       // Update validation flag in DB
       "DB_Recipes".Active_Recipe.Recipe_Valid := #Recipe_Valid;
       #Operation_OK := TRUE;
   END_IF;
END_FUNCTION

FUNCTION "FC_Safety_Monitor" : Void   // FC6, SCL
{ S7_Optimized_Access := 'TRUE' }
VERSION : 0.1
   VAR_INPUT
      Emergency_Stop : Bool;
      Door_Interlock_OK : Bool;
      Door_Locked : Bool;
      Manhole_Secured : Bool;
      Temperature_Value : Real;
      Pressure_Value : Real;
      System_Enabled : Bool;
   END_VAR
   VAR_OUTPUT
      Safety_OK : Bool;
      System_Ready : Bool;
      Emergency_Active : Bool;
      Safety_Fault : Bool;
      Fault_Code : UInt;
      Fault_Text : String;
   END_VAR
   VAR_TEMP
      Temp_High_Limit : Real;
      Pressure_High_Limit : Real;
   END_VAR
BEGIN
   #Safety_OK := TRUE;
   #Safety_Fault := FALSE;
   #Fault_Text := '';
   IF #Emergency_Stop THEN
       #Safety_OK := FALSE;
       #Safety_Fault := TRUE;
       #Fault_Text := 'EMERGENCY STOP ACTIVE';
       #System_Ready := FALSE;
       RETURN;
   END_IF;
   IF NOT #Door_Interlock_OK THEN
       #Safety_OK := FALSE;
       #Safety_Fault := TRUE;
       #Fault_Text := 'Door interlock not OK';
   END_IF;
   IF #Temperature_Value > 105.0 THEN
       #Safety_OK := FALSE;
       #Safety_Fault := TRUE;
       #Fault_Text := 'Temperature too high';
   END_IF;
   IF #Pressure_Value > 2500.0 THEN
       #Safety_OK := FALSE;
       #Safety_Fault := TRUE;
       #Fault_Text := 'Pressure too high';
   END_IF;
   #System_Ready := #Safety_OK AND #System_Enabled;
   IF #Safety_OK THEN
       #Fault_Text := 'All safety systems OK';
   END_IF;
END_FUNCTION

FUNCTION "FC_Lock_Discharge_Door" : Void   // FC7, SCL
{ S7_Optimized_Access := 'TRUE' }
VERSION : 0.1
   VAR_INPUT
      Step_Enable : Bool;
      Safety_OK : Bool;
      Step_Timeout : Time;
      Door_Locked_FB : Bool;
      Reset_Step : Bool;
   END_VAR
   VAR_OUTPUT
      Step_Complete : Bool;
      Step_Active : Bool;
      Step_Fault : Bool;
      Fault_Code : UInt;
      Status_Text : String;   // // Step status description
      Time_Remaining : Time;
   END_VAR
   VAR_IN_OUT
      Step_Timer : TON_TIME;
      Close_Timer : TON_TIME;
   END_VAR
BEGIN
   IF #Reset_Step THEN
       #Step_Timer(IN := FALSE,
                   PT := T#0S);
       #Step_Complete := FALSE;
       #Step_Active := FALSE;
       #Step_Fault := FALSE;
       #Fault_Code := 0;
       #Status_Text := 'Step reset';
       "DB_Valves".Valves[3].Close_Auto := FALSE;      // V3 discharge unlock
       RETURN;
   END_IF;
   IF #Step_Enable AND #Safety_OK THEN
       #Step_Active := TRUE;
       #Status_Text := 'Locking discharge door';

       "DB_Valves".Valves[3].Close_Auto := TRUE;       // V3 discharge unlock - close to
       #Step_Timer(IN := TRUE,
                   PT := #Step_Timeout);
       #Time_Remaining := #Step_Timeout - #Step_Timer.ET;
       #Close_Timer(IN := #Door_Locked_FB,
                    PT := T#2s);



       IF #Close_Timer.Q THEN
           #Step_Complete := TRUE;
           #Step_Active := FALSE;
           #Status_Text := 'Door locked successfully';
           "DB_Valves".Valves[3].Close_Auto := FALSE;

       ELSIF #Step_Timer.Q THEN
           #Step_Complete := FALSE;
           #Step_Active := FALSE;
           #Step_Fault := TRUE;
           #Fault_Code := 15;
           #Status_Text := 'Door lock timeout';
       END_IF;
   ELSE
       #Step_Active := FALSE;
       #Step_Complete := FALSE;
       #Step_Timer(IN := FALSE,
                   PT := T#0S);
       "DB_Valves".Valves[3].Close_Auto := FALSE;
       #Status_Text := 'Step disabled';
   END_IF;
END_FUNCTION

FUNCTION "FC_Add_Water" : Void   // FC8, SCL
{ S7_Optimized_Access := 'TRUE' }
VERSION : 0.1
   VAR_INPUT
      Step_Enable : Bool;
      Safety_OK : Bool;
      Reset_Step : Bool;
      Step_Timeout : Time;
      Target_Quantity : Real;
      Flow_Rate : Real;
   END_VAR
   VAR_OUTPUT
      Step_Complete : Bool;
      Water_Level_FB : Bool;
      Step_Active : Bool;
      Step_Fault : Bool;
      Fault_Code : UInt;
      Status_Text : String;
      Water_Added : Real;
      Time_Remaining : Time;
   END_VAR
   VAR_IN_OUT
      Step_Timer : TON_TIME;
   END_VAR
BEGIN
   IF #Reset_Step THEN
       #Step_Timer(IN := FALSE,
                   PT := T#0S);
       #Step_Complete := FALSE;
       #Step_Active := FALSE;
       #Step_Fault := FALSE;
       #Status_Text := 'Step reset';
       "DB_Valves".Valves[5].Open_Auto := FALSE;       // V5 water
       "DB_Valves".Valves[7].Open_Auto := FALSE;       // V7 evacuation
       #Water_Added := 0.0;
       RETURN;
   END_IF;

   IF #Step_Enable AND #Safety_OK THEN
       #Step_Active := TRUE;
       #Status_Text := 'Adding water';

       "DB_Valves".Valves[5].Open_Auto := TRUE;        // V5 water
       "DB_Valves".Valves[7].Open_Auto := TRUE;        // V7 evacuation
       "DB_Valves".Valves[3].Close_Auto := TRUE;         //V3
       #Step_Timer(IN := TRUE,
                   PT := #Step_Timeout);
       #Time_Remaining := #Step_Timeout - #Step_Timer.ET;

       IF #Flow_Rate > 0.0 THEN
           #Water_Added := (DINT_TO_REAL(TIME_TO_DINT(#Step_Timer.ET)) / 10.0) * #Flow_Rate;
           IF "DB_Recipes".Active_Recipe.Production.Adding_Water1_QTY < #Water_Added THEN
               "DB_Process".IO.Water_Level_FB := TRUE;
           END_IF;
       END_IF;

       IF "DB_Process".IO.Water_Level_FB THEN
           #Step_Complete := TRUE;
           #Step_Active := FALSE;
           #Status_Text := 'Water level reached';
           "DB_Valves".Valves[5].Open_Auto := FALSE;
       ELSIF #Step_Timer.Q THEN
           #Step_Complete := FALSE;
           #Step_Active := FALSE;
           #Step_Fault := TRUE;
           #Fault_Code := 1;
           #Status_Text := 'Water addition timeout';
       END_IF;
   ELSE
       #Step_Active := FALSE;
       #Step_Complete := FALSE;
       #Step_Timer(IN := FALSE,
                   PT := T#0S);
       "DB_Valves".Valves[5].Open_Auto := FALSE;
       "DB_Valves".Valves[7].Open_Auto := FALSE;
       #Status_Text := 'Step disabled';
   END_IF;
END_FUNCTION

FUNCTION "FC_Open_Manhole" : Void   // FC9, SCL
{ S7_Optimized_Access := 'TRUE' }
VERSION : 0.1
   VAR_INPUT
      Step_Enable : Bool;
      Safety_OK : Bool;
      Manhole_Open_FB : Bool;
      Manhole_Closed_FB : Bool;
      Reset_Step : Bool;
      Step_Timeout : Time;
   END_VAR
   VAR_OUTPUT
      Step_Complete : Bool;
      Step_Active : Bool;
      Step_Fault : Bool;
      Fault_Code : UInt;
      Status_Text : String;
      Time_Remaining : Time;   // // Time remaining in step
   END_VAR
   VAR_IN_OUT
      Step_Timer : TON_TIME;
      Open_Timer : TON_TIME;
   END_VAR
BEGIN
   IF #Reset_Step THEN
       #Step_Timer(IN := FALSE,
                   PT := T#0S);
       #Step_Complete := FALSE;
       #Step_Active := FALSE;
       #Step_Fault := FALSE;
       #Status_Text := 'Step reset';
       "DB_Valves".Valves[3].Open_Auto := FALSE;
       "DB_Valves".Valves[1].Open_Auto := FALSE;       // V1 manhole
       RETURN;
   END_IF;
   IF #Step_Enable AND #Safety_OK THEN
       #Step_Active := TRUE;
       #Status_Text := 'Opening manhole';

       "DB_Valves".Valves[1].Open_Auto := TRUE;        // V1 manhole
       "DB_Valves".Valves[3].Open_Auto := TRUE; 
       #Step_Timer(IN := TRUE,
                   PT := #Step_Timeout);
       #Time_Remaining := #Step_Timeout - #Step_Timer.ET;
       #Open_Timer(IN:=#Manhole_Closed_FB,
                   PT:=T#2S);
       IF #Open_Timer.Q THEN
           #Step_Complete := TRUE;
           #Step_Active := FALSE;
           #Status_Text := 'Manhole opened';
       ELSIF #Step_Timer.Q THEN
           #Step_Complete := FALSE;
           #Step_Active := FALSE;
           #Step_Fault := TRUE;
           #Fault_Code := 2;
           #Status_Text := 'Manhole open timeout';
       END_IF;
   ELSE
       #Step_Active := FALSE;
       #Step_Complete := FALSE;
       #Step_Timer(IN := FALSE,
                   PT := T#0S);
       "DB_Valves".Valves[1].Open_Auto := FALSE;
       "DB_Valves".Valves[3].Open_Auto := FALSE;
       #Status_Text := 'Step disabled';
   END_IF;
END_FUNCTION

FUNCTION "FC_Wait_Raw_Materials" : Void   // FC10, SCL
{ S7_Optimized_Access := 'TRUE' }
VERSION : 0.1
   VAR_INPUT
      Step_Enable : Bool;
      Safety_OK : Bool;
      RawMat_Confirm : Bool;   // // Raw materials loaded confirmation
      Manhole_Open_FB : Bool;   // // Manhole open feedback
      Manhole_Closed_FB : Bool;
      Reset_Step : Bool;
      Max_Wait_Time : Time;   // // Maximum wait time
   END_VAR
   VAR_OUTPUT
      Step_Complete : Bool;
      Step_Active : Bool;
      Step_Fault : Bool;
      Fault_Code : UInt;
      Status_Text : String;
      Wait_Time_Elapsed : Time;
   END_VAR
   VAR_IN_OUT
      Wait_Timer : TON_TIME;
   END_VAR
BEGIN
   IF #Reset_Step THEN
       #Wait_Timer(IN := FALSE,
                   PT := T#0S);
       #Step_Complete := FALSE;
       #Step_Active := FALSE;
       #Step_Fault := FALSE;
       #Status_Text := 'Step reset';
       RETURN;
   END_IF;
   IF #Step_Enable AND #Safety_OK THEN
       #Step_Active := TRUE;
       #Status_Text := 'Waiting for raw materials';

       "DB_Valves".Valves[1].Open_Auto := TRUE;        // V1 manhole - keep open
       "DB_Valves".Valves[3].Open_Auto := TRUE;        // V7 evacuation
       #Wait_Timer(IN := TRUE,
                   PT := #Max_Wait_Time);
       #Wait_Time_Elapsed := #Wait_Timer.ET;

       IF  #Manhole_Closed_FB THEN
           #Step_Complete := FALSE;
           #Step_Active := FALSE;
           #Step_Fault := TRUE;
           #Fault_Code := 3;
           #Status_Text := 'Manhole not open-Reset PLS';
           RETURN;
       END_IF;

       IF #RawMat_Confirm THEN
           #Step_Complete := TRUE;
           #Step_Active := FALSE;
           #Status_Text := 'Raw materials confirmed';
       ELSIF #Wait_Timer.Q THEN
           #Status_Text := 'Long wait time - check operator';
           #Wait_Timer(IN := FALSE,
                       PT := T#0S);
       END_IF;
   ELSE
       #Step_Active := FALSE;
       #Step_Complete := FALSE;
       #Wait_Timer(IN := FALSE,
                   PT := T#0S);
       #Status_Text := 'Step disabled';
   END_IF;
END_FUNCTION

FUNCTION "FC_Close_Manhole" : Void   // FC11, SCL
{ S7_Optimized_Access := 'TRUE' }
VERSION : 0.1
   VAR_INPUT
      Step_Enable : Bool;
      Safety_OK : Bool;
      Step_Timeout : Time;
      Manhole_Closed_FB : Bool;
      Reset_Step : Bool;
      Manhole_Open_FB : Bool;
   END_VAR
   VAR_OUTPUT
      Step_Complete : Bool;
      Step_Active : Bool;
      Step_Fault : Bool;
      Fault_Code : UInt;
      Status_Text : String;
      Time_Remaining : Time;
   END_VAR
   VAR_IN_OUT
      Step_Timer : TON_TIME;
      Close_Timer : TON_TIME;
   END_VAR
BEGIN
   IF #Reset_Step THEN
       #Step_Timer(IN := FALSE,
                   PT := T#0S);
       #Step_Complete := FALSE;
       #Step_Active := FALSE;
       #Step_Fault := FALSE;
       #Status_Text := 'Step reset';
       "DB_Valves".Valves[1].Close_Auto := FALSE;      // V1 manhole
       "DB_Valves".Valves[3].Close_Auto := FALSE;
       "DB_Valves".Valves[2].Open_Auto := FALSE;

       RETURN;
   END_IF;
   IF #Step_Enable AND #Safety_OK THEN
       #Step_Active := TRUE;
       #Status_Text := 'Closing manhole';

       "DB_Valves".Valves[1].Open_Auto := FALSE;       // V1 manhole - stop opening
       "DB_Valves".Valves[1].Close_Auto := TRUE;       // V1 manhole - start closing
       "DB_Valves".Valves[3].Close_Auto := TRUE;
       "DB_Valves".Valves[2].Open_Auto := TRUE;
       #Step_Timer(IN := TRUE,
                   PT := #Step_Timeout);
       #Time_Remaining := #Step_Timeout - #Step_Timer.ET;
       #Close_Timer(IN := #Manhole_Closed_FB,
                    PT := t#2s);
       IF #Close_Timer.Q THEN
           #Step_Complete := TRUE;
           #Step_Active := FALSE;
           #Status_Text := 'Manhole closed & secured';
           "DB_Valves".Valves[1].Close_Auto := FALSE;
       ELSIF #Step_Timer.Q THEN
           #Step_Complete := FALSE;

           #Step_Active := FALSE;
           #Step_Fault := TRUE;
           #Fault_Code := 4;
           #Status_Text := 'Manhole close timeout';
       END_IF;
   ELSE
       #Step_Active := FALSE;
       #Step_Complete := FALSE;
       #Step_Timer(IN := FALSE,
                   PT := T#0S);
       "DB_Valves".Valves[1].Open_Auto := FALSE;
       "DB_Valves".Valves[1].Close_Auto := FALSE;
       "DB_Valves".Valves[3].Close_Auto := FALSE;
       "DB_Valves".Valves[2].Open_Auto := FALSE;
       #Status_Text := 'Step disabled';
   END_IF;
END_FUNCTION

FUNCTION "FC_Valve_Integration" : Void   // FC12, SCL
{ S7_Optimized_Access := 'TRUE' }
VERSION : 0.1
   VAR_INPUT
      Valve_Number : UInt;
   END_VAR
   VAR_OUTPUT
      Integration_OK : Bool;
   END_VAR
   VAR_IN_OUT
      Valve_Data : "UDT_Valve";
      Valve_FB_Instance : "FB_Valve_DO";
   END_VAR
BEGIN
   // Set valve name based on number
   CASE #Valve_Number OF
       1:
           #Valve_Data.Config.Valve_Name := 'V1_MANHOLE';
       2:
           #Valve_Data.Config.Valve_Name := 'V2_CIP';
       3:
           #Valve_Data.Config.Valve_Name := 'V3_DISCHARGE_UNLOCK';
       4:
           #Valve_Data.Config.Valve_Name := 'V4_DISCHARGE_OPEN';
       5:
           #Valve_Data.Config.Valve_Name := 'V5_WATER_SUPPLY';
       6:
           #Valve_Data.Config.Valve_Name := 'V6_STEAM';
       7:
           #Valve_Data.Config.Valve_Name := 'V7_EVACUATION';
       8:
           #Valve_Data.Config.Valve_Name := 'V8_VACUUM';
       9:
           #Valve_Data.Config.Valve_Name := 'V9_VACUUM_COOLING';
   END_CASE;

   // Map UDT commands to your FB inputs  
   #Valve_FB_Instance(
                      // Command inputs
                      AutoCmd := #Valve_Data.Command.Open_Auto,
                      FuncCmd := #Valve_Data.Command.Open_Func,
                      ManCmd := #Valve_Data.Command.Open_Man,
                      OOS := #Valve_Data.Interlocks.OOS,
                      Permissive := #Valve_Data.Interlocks.Permissive,
                      FbOpen := #Valve_Data.Status.Limit_Open,
                      FbClosed := #Valve_Data.Status.Limit_Closed,
                      TwoCoils := #Valve_Data.Config.TwoCoils,
                      T_Stroke := #Valve_Data.Config.Stroke_Time,
                      T_Timeout := #Valve_Data.Config.Travel_Timeout,

                      // Output mappings
                      Q_Open => #Valve_Data.Outputs.Q_Run,
                      Q_Close => #Valve_Data.Outputs.Q_Close,
                      Ready => #Valve_Data.Status.Ready,
                      FaultTO => #Valve_Data.Status.Fault,
                      FaultFB => #Valve_Data.Status.Fault,
                      Source => #Valve_Data.Status.Source,
                      Status => #Valve_Data.Status.State
   );

   // Update valve status based on FB outputs
   IF #Valve_Data.Status.Limit_Open THEN
       #Valve_Data.Status.State := 3;      // Open
   ELSIF #Valve_Data.Status.Limit_Closed THEN
       #Valve_Data.Status.State := 1;      // Closed
   ELSIF #Valve_Data.Outputs.Q_Run THEN
       #Valve_Data.Status.State := 2;      // Opening
   ELSIF #Valve_Data.Outputs.Q_Close THEN
       #Valve_Data.Status.State := 4;      // Closing  
   ELSE
       #Valve_Data.Status.State := 0;      // Unknown
   END_IF;

   #Integration_OK := TRUE;
END_FUNCTION

ORGANIZATION_BLOCK "Main"   // OB1, LAD, ProgramCycle
TITLE = "Main Program Sweep (Cycle)"
{ S7_Optimized_Access := 'TRUE' }
VERSION : 0.1
   VAR_INPUT
      Initial_Call : Bool;   // Initial call of this OB
      Remanence : Bool;   // =True, if remanent data are available
   END_VAR
   VAR_TEMP
      TempOffset : Bool;
      Temp_DINT : DInt;
      First_Scan : Bool;
   END_VAR
BEGIN

REGION Network 1: First Scan & Process Main FB Call
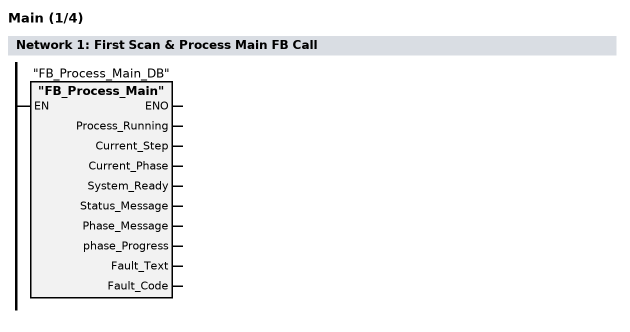
   RUNG wire#powerrail
      "FB_Process_Main_DB"(Process_Running =>, Current_Step =>, Current_Phase =>, System_Ready =>, Status_Message =>, Phase_Message =>, phase_Progress =>, Fault_Text =>, Fault_Code =>)
   END_RUNG
   // the same network as SCL:
   "FB_Process_Main_DB"();   // "FB_Process_Main"
END_REGION

REGION Network 2: Alarms
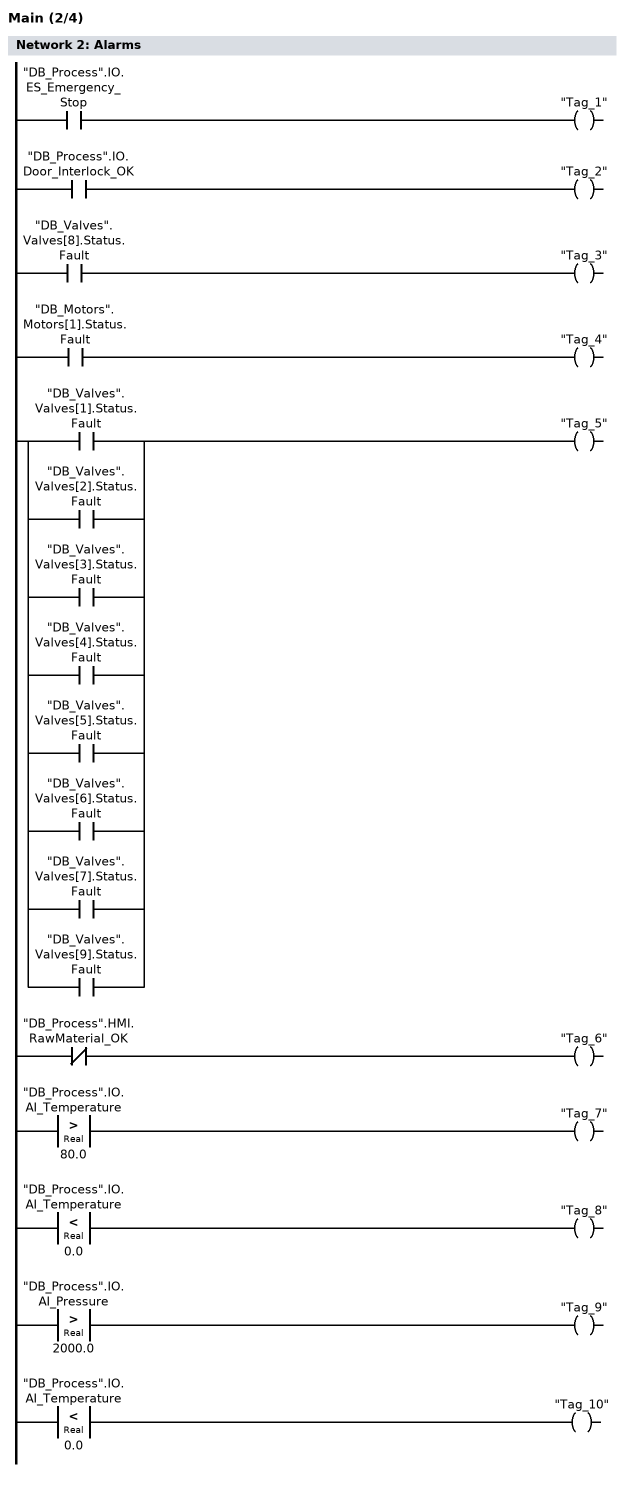
   RUNG wire#powerrail
      Contact( "DB_Process".IO.ES_Emergency_Stop )
      Coil( "Tag_1" )
   END_RUNG
   RUNG wire#powerrail
      Contact( "DB_Process".IO.Door_Interlock_OK )
      Coil( "Tag_2" )
   END_RUNG
   RUNG wire#powerrail
      Contact( "DB_Valves".Valves[8].Status.Fault )
      Coil( "Tag_3" )
   END_RUNG
   RUNG wire#powerrail
      Contact( "DB_Motors".Motors[1].Status.Fault )
      Coil( "Tag_4" )
   END_RUNG
   RUNG wire#powerrail
      Contact( "DB_Valves".Valves[1].Status.Fault )
      wire#w1
      Coil( "Tag_5" )
   END_RUNG
   RUNG wire#powerrail
      Contact( "DB_Valves".Valves[2].Status.Fault )
   END_RUNG wire#w1
   RUNG wire#powerrail
      Contact( "DB_Valves".Valves[3].Status.Fault )
   END_RUNG wire#w1
   RUNG wire#powerrail
      Contact( "DB_Valves".Valves[4].Status.Fault )
   END_RUNG wire#w1
   RUNG wire#powerrail
      Contact( "DB_Valves".Valves[5].Status.Fault )
   END_RUNG wire#w1
   RUNG wire#powerrail
      Contact( "DB_Valves".Valves[6].Status.Fault )
   END_RUNG wire#w1
   RUNG wire#powerrail
      Contact( "DB_Valves".Valves[7].Status.Fault )
   END_RUNG wire#w1
   RUNG wire#powerrail
      Contact( "DB_Valves".Valves[9].Status.Fault )
   END_RUNG wire#w1
   RUNG wire#powerrail
      I_Contact( "DB_Process".HMI.RawMaterial_OK )
      Coil( "Tag_6" )
   END_RUNG
   RUNG wire#powerrail
      { S7_Templates := "SrcType := Real" } GT_Contact(in1 := "DB_Process".IO.AI_Temperature, in2 := 80.0)
      Coil( "Tag_7" )
   END_RUNG
   RUNG wire#powerrail
      { S7_Templates := "SrcType := Real" } LT_Contact(in1 := "DB_Process".IO.AI_Temperature, in2 := 0.0)
      Coil( "Tag_8" )
   END_RUNG
   RUNG wire#powerrail
      { S7_Templates := "SrcType := Real" } GT_Contact(in1 := "DB_Process".IO.AI_Pressure, in2 := 2000.0)
      Coil( "Tag_9" )
   END_RUNG
   RUNG wire#powerrail
      { S7_Templates := "SrcType := Real" } LT_Contact(in1 := "DB_Process".IO.AI_Temperature, in2 := 0.0)
      Coil( "Tag_10" )
   END_RUNG
   // the same network as SCL:
   "Tag_1" := "DB_Process".IO.ES_Emergency_Stop;
   "Tag_2" := "DB_Process".IO.Door_Interlock_OK;
   "Tag_3" := "DB_Valves".Valves[8].Status.Fault;
   "Tag_4" := "DB_Motors".Motors[1].Status.Fault;
   "Tag_5" := "DB_Valves".Valves[1].Status.Fault OR "DB_Valves".Valves[2].Status.Fault OR "DB_Valves".Valves[3].Status.Fault OR "DB_Valves".Valves[4].Status.Fault OR "DB_Valves".Valves[5].Status.Fault OR "DB_Valves".Valves[6].Status.Fault OR "DB_Valves".Valves[7].Status.Fault OR "DB_Valves".Valves[9].Status.Fault;
   "Tag_6" := NOT "DB_Process".HMI.RawMaterial_OK;
   "Tag_7" := "DB_Process".IO.AI_Temperature > 80.0;
   "Tag_8" := "DB_Process".IO.AI_Temperature < 0.0;
   "Tag_9" := "DB_Process".IO.AI_Pressure > 2000.0;
   "Tag_10" := "DB_Process".IO.AI_Temperature < 0.0;
END_REGION

REGION Network 3: Digital Input Mapping
   // "DB_Process".IO.Door_Locked_FB , "DB_Process".IO.Manhole_Closed_FB, "DB_Process".IO.Manhole_Open_FB, "DB_Process".IO.Water_Level_FB, "DB_Process".IO.Door_Interlock_OK, "DB_Process".IO.ES_Emergency_Stop
END_REGION

REGION Network 4: "Analog Input - Temperature Scaling"
END_REGION

REGION Network 5: "Analog Input - Pressure Scaling"
   // "Pressure Input", water flow
END_REGION

REGION Network 6: Analog Input Scaling - Water Flow
END_REGION

REGION Network 7: Digital Output Mapping - Motor
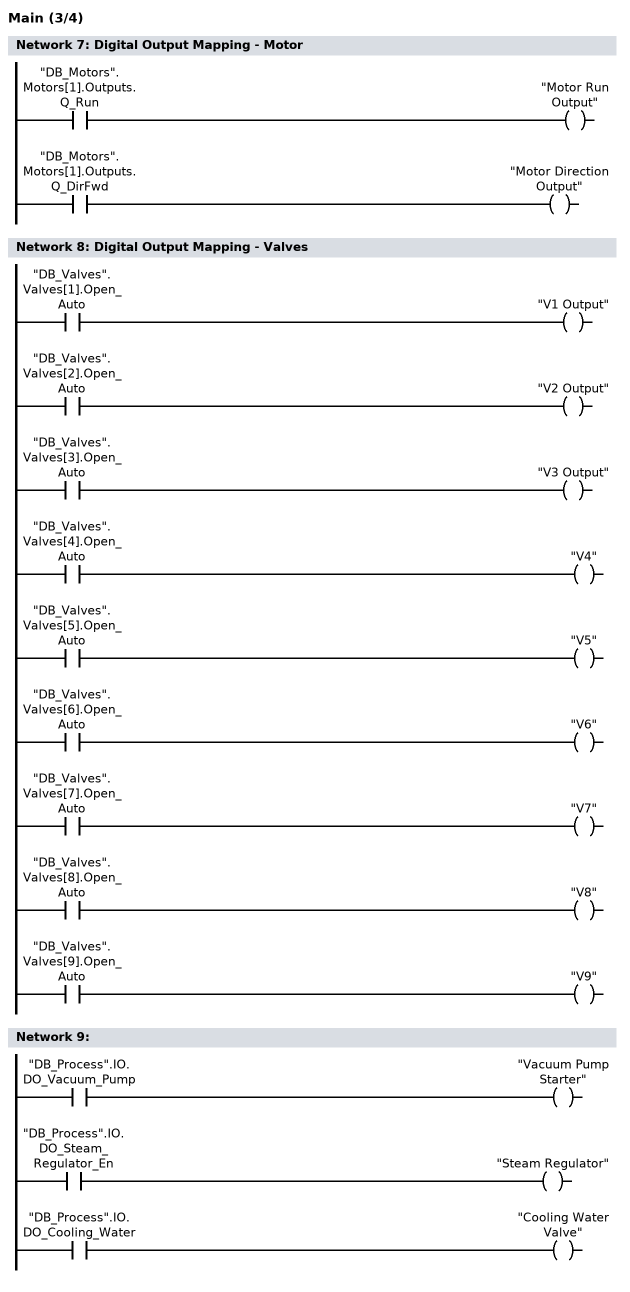
   RUNG wire#powerrail
      Contact( "DB_Motors".Motors[1].Outputs.Q_Run )
      Coil( "Motor Run Output" )
   END_RUNG
   RUNG wire#powerrail
      Contact( "DB_Motors".Motors[1].Outputs.Q_DirFwd )
      Coil( "Motor Direction Output" )
   END_RUNG
   // the same network as SCL:
   "Motor Run Output" := "DB_Motors".Motors[1].Outputs.Q_Run;
   "Motor Direction Output" := "DB_Motors".Motors[1].Outputs.Q_DirFwd;
END_REGION

REGION Network 8: Digital Output Mapping - Valves
   RUNG wire#powerrail
      Contact( "DB_Valves".Valves[1].Open_Auto )
      Coil( "V1 Output" )
   END_RUNG
   RUNG wire#powerrail
      Contact( "DB_Valves".Valves[2].Open_Auto )
      Coil( "V2 Output" )
   END_RUNG
   RUNG wire#powerrail
      Contact( "DB_Valves".Valves[3].Open_Auto )
      Coil( "V3 Output" )
   END_RUNG
   RUNG wire#powerrail
      Contact( "DB_Valves".Valves[4].Open_Auto )
      Coil( "V4" )
   END_RUNG
   RUNG wire#powerrail
      Contact( "DB_Valves".Valves[5].Open_Auto )
      Coil( "V5" )
   END_RUNG
   RUNG wire#powerrail
      Contact( "DB_Valves".Valves[6].Open_Auto )
      Coil( "V6" )
   END_RUNG
   RUNG wire#powerrail
      Contact( "DB_Valves".Valves[7].Open_Auto )
      Coil( "V7" )
   END_RUNG
   RUNG wire#powerrail
      Contact( "DB_Valves".Valves[8].Open_Auto )
      Coil( "V8" )
   END_RUNG
   RUNG wire#powerrail
      Contact( "DB_Valves".Valves[9].Open_Auto )
      Coil( "V9" )
   END_RUNG
   // the same network as SCL:
   "V1 Output" := "DB_Valves".Valves[1].Open_Auto;
   "V2 Output" := "DB_Valves".Valves[2].Open_Auto;
   "V3 Output" := "DB_Valves".Valves[3].Open_Auto;
   "V4" := "DB_Valves".Valves[4].Open_Auto;
   "V5" := "DB_Valves".Valves[5].Open_Auto;
   "V6" := "DB_Valves".Valves[6].Open_Auto;
   "V7" := "DB_Valves".Valves[7].Open_Auto;
   "V8" := "DB_Valves".Valves[8].Open_Auto;
   "V9" := "DB_Valves".Valves[9].Open_Auto;
END_REGION

REGION Network 9
   RUNG wire#powerrail
      Contact( "DB_Process".IO.DO_Vacuum_Pump )
      Coil( "Vacuum Pump Starter" )
   END_RUNG
   RUNG wire#powerrail
      Contact( "DB_Process".IO.DO_Steam_Regulator_En )
      Coil( "Steam Regulator" )
   END_RUNG
   RUNG wire#powerrail
      Contact( "DB_Process".IO.DO_Cooling_Water )
      Coil( "Cooling Water Valve" )
   END_RUNG
   // the same network as SCL:
   "Vacuum Pump Starter" := "DB_Process".IO.DO_Vacuum_Pump;
   "Steam Regulator" := "DB_Process".IO.DO_Steam_Regulator_En;
   "Cooling Water Valve" := "DB_Process".IO.DO_Cooling_Water;
END_REGION

REGION Network 10
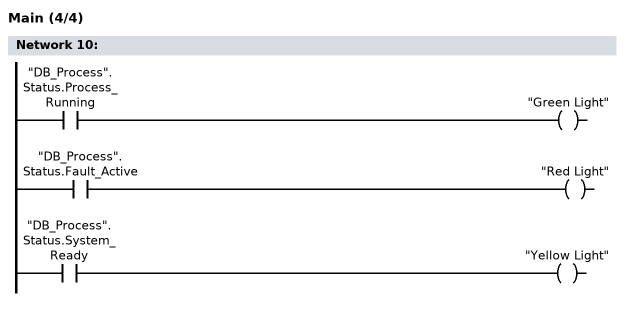
   RUNG wire#powerrail
      Contact( "DB_Process".Status.Process_Running )
      Coil( "Green Light" )
   END_RUNG
   RUNG wire#powerrail
      Contact( "DB_Process".Status.Fault_Active )
      Coil( "Red Light" )
   END_RUNG
   RUNG wire#powerrail
      Contact( "DB_Process".Status.System_Ready )
      Coil( "Yellow Light" )
   END_RUNG
   // the same network as SCL:
   "Green Light" := "DB_Process".Status.Process_Running;
   "Red Light" := "DB_Process".Status.Fault_Active;
   "Yellow Light" := "DB_Process".Status.System_Ready;
END_REGION
END_ORGANIZATION_BLOCK

(* ===== HMI "HMI_RT_2" =====
system functions are stored by id; their names below are inferred from use
connection "HMI_Connection_2": ETHERNET, S7_1200_OMS

HMI tags "Default tag table"
   "Tag_ScreenNumber" : UInt, internal
   "HMI_Alarm_Word" : Int = PLC DB_Process.Status.Current_Step AT %MW3, 1 s
   "DB_Motors_Motors{1}_Config_Max_Speed_pct" : Real = PLC DB_Process.Status.Current_Phase, 1 s
   "DB_Motors_Motors{1}_Config_Min_Speed_pct" : Real = PLC DB_Process.Status.Process_Running, 1 s
   "Manhole_open_FB" : Bool = PLC DB_Process.Status.System_Ready AT %DB21.DBX875.6, 1 s
   "Water_level" : Real = PLC DB_Process.Status.Water_Level_Actual AT %DB21.DBD554, 1 s
   "Door_interlock" : Bool = PLC DB_Process.IO.Door_Interlock_OK AT %DB21.DBX875.1, 1 s

HMI tags "Process Status Tags"
   "HMI_Current_Step" : UInt = PLC DB_Process.Status.Current_Step AT %DB21.DBW0, 1 s
   "HMI_Current_Phase" : UInt = PLC DB_Process.Status.Current_Phase AT %DB21.DBW516, 1 s
   "HMI_Process_Running" : Bool = PLC DB_Process.Status.Process_Running AT %DB21.DBX574.0, 1 s
   "HMI_System_Ready" : Bool = PLC DB_Process.Status.System_Ready AT %DB21.DBX574.7, 1 s
   "HMI_Progress" : Real = PLC FB_Process_Main_DB.phase_Progress AT %DB21.DBD274, 1 s
   "HMI_Status_Message" : String[254] = PLC DB_Process.Status.Step_Name AT %DB21.DBX2.0, 1 s
   "HMI_Individual_Discharg" : Bool = PLC DB_Process.Status.Individual_Discharge_Active AT %DB21.DBX580.0, 100 ms
   "Phase_Message" : String[254] = PLC DB_Process.Status.Phase_Name AT %DB21.DBX258.0, 1 s

HMI tags "Process Values Tags"
   "HMI_Temperature" : Real = PLC DB_Process.IO.AI_Temperature AT %DB21.DBD876, 1 s
   "HMI_Pressure" : Real = PLC DB_Process.IO.AI_Pressure AT %DB21.DBD880, 1 s
   "HMI_Water_Flow" : Real = PLC DB_Process.IO.AI_Water_Flow AT %DB21.DBD888, 1 s
   "HMI_Motor_Speed" : Real = PLC DB_Motors.Motors[1].Outputs.AO_SpeedPct, 1 s
   "HMI_Steam_Position" : Real = PLC DB_Process.IO.AO_Steam_Regulator AT %DB21.DBD910, 1 s
   "Cooking Time" : Time = PLC DB_Recipes.Active_Recipe.Production.Cooking_Time_Phase1 AT %DB1.DBD0, 1 s
   "Cold Mix Time" : Time = PLC DB_Recipes.Active_Recipe.Production.Cold_Mix_Time AT %DB1.DBD0, 1 s
   "Forward Time" : Time = PLC FB_Motor_VFD_DB.Tmr_Fwd.PT AT %DB1.DBD0, 1 s
   "FB_Motor_VFD_DB_Tmr_Bwd_PT" : Time = PLC FB_Motor_VFD_DB.Tmr_Bwd.PT AT %DB1.DBD0, 1 s
   "Vaccum Setpoint" : Real = PLC DB_Recipes.Active_Recipe.Vacuum.Vacuum_Setpoint_mbar AT %DB1.DBD0, 1 s
   "Water Quant." : Real = PLC DB_Recipes.Active_Recipe.Production.Adding_Water1_QTY AT %DB1.DBD0, 1 s

HMI tags "Equipment Status Tags"
   "HMI_Motor_Running" : Bool = PLC DB_Motors.Motors[1].Status.Running, 500 ms
   "HMI_V1_Open" : Bool = PLC DB_Valves.Valves[1].Open_Auto AT %DB1.DBW0, 500 ms
   "HMI_V1_Closed" : Bool = PLC DB_Valves.Valves[1].Close_Auto AT %DB1.DBW0, 500 ms
   "HMI_V3_Open" : Bool = PLC DB_Valves.Valves[3].Open_Auto AT %DB1.DBW0, 500 ms
   "HMI_V4_Open" : Bool = PLC DB_Valves.Valves[4].Open_Auto AT %DB1.DBW0, 500 ms
   "HMI_V5_Open" : Bool = PLC DB_Valves.Valves[5].Open_Auto AT %DB1.DBW0, 500 ms
   "HMI_V6_Open" : Bool = PLC DB_Valves.Valves[6].Open_Auto AT %DB1.DBW0, 500 ms
   "HMI_V7_Open" : Bool = PLC DB_Valves.Valves[7].Open_Auto AT %DB1.DBW0, 500 ms
   "HMI_V8_Open" : Bool = PLC DB_Valves.Valves[8].Open_Auto AT %DB1.DBW0, 500 ms
   "HMI_V9_Open" : Bool = PLC DB_Valves.Valves[9].Status.Open AT %DB1.DBW0, 500 ms
   "HMI_Door_Locked" : Bool = PLC DB_Process.IO.Door_Locked_FB AT %DB21.DBX875.3, 500 ms
   "HMI_Manhole_Closed" : Bool = PLC DB_Process.IO.Manhole_Closed_FB AT %DB21.DBX875.7, 500 ms
   "HMI_V1_Fault" : Bool = PLC DB_Valves.Valves[1].Status.Fault AT %DB1.DBX0.0, 1 s
   "HMI_V2_Fault" : Bool = PLC DB_Valves.Valves[2].Status.Fault AT %DB1.DBX0.0, 1 s
   "HMI_V3_Fault" : Bool = PLC DB_Valves.Valves[3].Status.Fault AT %DB1.DBX0.0, 1 s
   "HMI_V4_Fault" : Bool = PLC DB_Valves.Valves[4].Status.Fault AT %DB1.DBX0.0, 1 s
   "HMI_V5_Fault" : Bool = PLC DB_Valves.Valves[5].Status.Fault AT %DB1.DBX0.0, 1 s
   "HMI_V6_Fault" : Bool = PLC DB_Valves.Valves[6].Status.Fault AT %DB1.DBX0.0, 1 s
   "HMI_V7_Fault" : Bool = PLC DB_Valves.Valves[7].Status.Fault AT %DB1.DBX0.0, 1 s
   "HMI_V8_Fault" : Bool = PLC DB_Valves.Valves[8].Status.Fault AT %DB1.DBX0.0, 1 s
   "HMI_V9_Fault" : Bool = PLC DB_Valves.Valves[9].Status.Fault AT %DB1.DBX0.0, 1 s
   "HMI_V2_Open" : Bool = PLC DB_Valves.Valves[2].Open_Auto AT %DB1.DBX0.0, 1 s
   "HMI_Direction" : UInt = PLC DB_Motors.Motors[1].Status.Direction AT %DB1.DBX0.0, 1 s
   "HMI_V3_close" : Bool = PLC DB_Valves.Valves[3].Close_Auto AT %DB1.DBX0.0, 1 s

HMI tags "Control Command Tags"
   "DB_Process_HMI_Start_Production" : Bool = PLC DB_Process.HMI.Start_Production AT %DB21.DBX582.0, 500 ms
   "HMI_Stop_Production" : Bool = PLC DB_Process.HMI.Stop_Production AT %DB21.DBX582.1, 500 ms
   "HMI_Reset_System" : Bool = PLC DB_Process.HMI.Reset_System AT %DB21.DBX582.2, 500 ms
   "HMI_Emergency_Stop" : Bool = PLC DB_Process.IO.ES_Emergency_Stop AT %DB21.DBX874.5, 100 ms
   "HMI_RawMaterial_OK" : Bool = PLC DB_Process.HMI.RawMaterial_OK AT %DB21.DBX582.6, 1 s
   "HMI_Discharge_Ready_OK" : Bool = PLC DB_Process.HMI.Discharge_Ready_OK AT %DB21.DBX583.0, 1 s
   "Green_Light HMI" : Bool = PLC "Green Light" AT %Q3.0, 1 s
   "Red light HMI" : Bool = PLC "Red Light" AT %Q3.2, 1 s
   "Yellow Light HMI" : Bool = PLC "Yellow Light" AT %Q3.1, 1 s
   "Reset_p_s" : Bool = PLC DB_Process.HMI.Reset_p_s AT %DB21.DBX582.3, 1 s
   "Direction Motor" : UInt = PLC DB_Motors.Motors[1].Status.State AT %DB1.DBX0.0, 1 s
   "water_LEVEL_FB" : Bool = PLC DB_Process.IO.Water_Level_FB AT %DB21.DBX875.5, 1 s
   "HMI_Acknowledge_Word" : Int = PLC Acknowledge_Word AT %MW4, 1 s
   "HMI_Acknowledge_bit" : Bool = PLC "Acknowledge bit" AT %M5.0, 1 s

HMI tags "Manual Control Tags"
   "HMI_V1_Manual_Open" : Bool = PLC DB_Valves.Valves[1].Open_Man AT %DB1.DBW0, 500 ms
   "HMI_V1_Manual_Close" : Bool = PLC DB_Valves.Valves[1].Close_Man AT %DB1.DBX0.0, 1 s
   "HMI_V2_Manual_Open" : Bool = PLC DB_Valves.Valves[2].Open_Man AT %DB1.DBW0, 500 ms
   "HMI_V2_Manual_Close" : Bool = PLC DB_Valves.Valves[2].Close_Man AT %DB1.DBX0.0, 1 s
   "HMI_V3_Manual_Open" : Bool = PLC DB_Valves.Valves[3].Open_Man AT %DB1.DBW0, 500 ms
   "HMI_V3_Manual_Close" : Bool = PLC DB_Valves.Valves[3].Close_Man AT %DB1.DBX0.0, 1 s
   "HMI_V4_Manual_Open" : Bool = PLC DB_Valves.Valves[4].Open_Man AT %DB1.DBW0, 500 ms
   "HMI_V4_Manual_Close" : Bool = PLC DB_Valves.Valves[4].Close_Man AT %DB1.DBX0.0, 1 s
   "HMI_V5_Manual_Open" : Bool = PLC DB_Valves.Valves[5].Open_Man AT %DB1.DBW0, 500 ms
   "HMI_V5_Manual_Close" : Bool = PLC DB_Valves.Valves[5].Close_Man AT %DB1.DBX0.0, 1 s
   "HMI_V6_Manual_Open" : Bool = PLC DB_Valves.Valves[6].Open_Man AT %DB1.DBW0, 500 ms
   "HMI_V6_Manual_Close" : Bool = PLC DB_Valves.Valves[6].Close_Man AT %DB1.DBX0.0, 1 s
   "HMI_V7_Manual_Open" : Bool = PLC DB_Valves.Valves[7].Open_Man AT %DB1.DBW0, 500 ms
   "HMI_V7_Manual_Close" : Bool = PLC DB_Valves.Valves[7].Close_Man AT %DB1.DBX0.0, 1 s
   "HMI_V8_Manual_Open" : Bool = PLC DB_Valves.Valves[8].Open_Man AT %DB1.DBW0, 500 ms
   "HMI_V8_Manual_Close" : Bool = PLC DB_Valves.Valves[8].Close_Man AT %DB1.DBX0.0, 1 s
   "HMI_V9_Manual_Open" : Bool = PLC DB_Valves.Valves[9].Open_Man AT %DB1.DBW0, 500 ms
   "HMI_V9_Manual_Close" : Bool = PLC DB_Valves.Valves[9].Close_Man AT %DB1.DBX0.0, 1 s
   "HMI_Motor_Manual_Start" : Bool = PLC DB_Motors.Motors[1].Command.Start_Man, 1 s
   "HMI_Motor_Manual_Stop" : Bool = PLC DB_Motors.Motors[1].Command.Stop, 1 s

discrete alarms
   1: 'Emergency stop activated', class Errors, trigger "HMI_Alarm_Word" bit 0
   2: 'Motor fault detected', class Errors, trigger "HMI_Alarm_Word" bit 7
   3: 'Vacuum system fault or deviation beyond tolerance', class Errors, trigger "HMI_Alarm_Word" bit 6
   4: 'Pressure below safe limits', class Errors, trigger "HMI_Alarm_Word" bit 5
   5: 'Steam pressure exceeds maximum safe pressure', class Errors, trigger "HMI_Alarm_Word" bit 4
   6: 'Product temperature below low alarm setpoint', class Errors, trigger "HMI_Alarm_Word" bit 3
   7: 'Product temperature exceeds high alarm setpoint', class Errors, trigger "HMI_Alarm_Word" bit 2
   8: 'Raw material loading step timeout or not confirmed', class Errors, trigger "HMI_Alarm_Word" bit 10
   9: 'Any system-wide fault or fault mask active', class Errors, trigger "HMI_Alarm_Word" bit 13
   11: 'Motor fault detected', class Errors, trigger "HMI_Alarm_Word" bit 8
   10: 'Interlock is activiated', class Warnings, trigger "HMI_Alarm_Word" bit 1

SlideinScreen "GraphX_Slidein_Left" 267x480
   TextField "Text field_11" at 0,246 size 117x23; Text 'Vacuum Set.'

screen "MAIN LAYOUT SCREEN" 800x420, template "Template_1"
   on GenerateScreen: SetTag("Tag_ScreenNumber", 1)
   GraphicView "Graphic view_1" at 547,303 size 57x46; Picture "Graphic_1"
   Button "Button_1" at 557,307 size 39x38; TextOff 'Text'
   SymbolLibrary "Symbol library_6" at -2,1 size 803x422
   Button "HmiScreenItemData" at 0,366 size 128x47; TextOff 'Parameters'; TextOn 'Sub Open/Close Manhole'; PictureOff "Navigates to Sub Open/Close Manhole for TP700 Comfort 17.0.0.0"; PictureOn "Navigates to Sub Open/Close Manhole for TP700 Comfort 17.0.0.0"
      on Press: function_efd93a16("parameters", 0, 0, -1, -1, 1)
   TextField "Text field_2" at 86,97 size 16x23; Text 'Text'
   Group "Group" at 547,303 size 57x46; Picture "Graphic_1"
   SymbolLibrary "Symbol library_1" at 231,207 size 57x44
   SymbolLibrary "Symbol library_3" at 334,89 size 343x244
      on Activate: function_efd93a16("motor manual", 0, 0, -1, -1, 1)
   IOField "I/O field_7" at 464,171 size 87x37; FormatPattern 9999
      ProcessValue <- "HMI_Motor_Speed"
   GraphicView "Graphic view_4" at 216,68 size 78x64; Picture "Graphic_7"
   SymbolLibrary "Symbol library_5" at 259,204 size 57x44
      Appearance <- "Water_level"
   SymbolLibrary "Symbol library_2" at 660,122 size 23x202
      on Press: InvertBit("HMI_Door_Locked")
      Visibility <- "HMI_Door_Locked"
   Polygon "Polygon_1" at 337,79 size 338x43
      Appearance <- "HMI_Manhole_Closed"
   TextField "Text field_11" at 487,89 size 66x20; Text 'Manhole'
   IOField "I/O field_4" at 82,187 size 96x38; FormatPattern s999999999.999
      ProcessValue <- "HMI_Temperature"
   TextField "Text field_7" at 83,164 size 100x20; Text 'Temperature'
   TextField "Text field_6" at 101,163 size 49x20; Text 'Phase'
   IOField "I/O field_3" at 102,183 size 47x38; FormatPattern 99
      ProcessValue <- "HMI_Current_Phase"
   TextField "Text field_4" at 89,98 size 82x28; Text 'Current Step'
   IOField "I/O field_1" at 100,119 size 47x38; FormatPattern 99
      ProcessValue <- "HMI_Current_Step"
   IOField "I/O field_2" at 0,28 size 185x33; FormatPattern ????????????????????????????????????????
      ProcessValue <- "Phase_Message"
   TextField "Text field_1" at 5,11 size 203x20; Text 'Production Status & Steps'
   IOField "I/O field_6" at 94,309 size 82x39; FormatPattern 9999
      ProcessValue <- "HMI_Water_Flow"
   TextField "Text field_10" at 95,287 size 88x20; Text 'Water Flow'
   SymbolLibrary "Symbol library_9" at 624,44 size 65x62
   SymbolLibrary "Symbol library_10" at 305,216 size 65x37
   SymbolLibrary "Symbol library_11" at 202,228 size 64x44
   SymbolLibrary "Symbol library_12" at 198,265 size 33x44
   SymbolLibrary "Symbol library_13" at 198,275 size 65x65
   SymbolLibrary "Symbol library_14" at 292,315 size 65x44
   SymbolLibrary "Symbol library_15" at 600,281 size 57x44
      on Press: InvertBit("Door_interlock")
      Appearance <- "Door_interlock"
   SymbolLibrary "Symbol library_16" at 597,144 size 57x44
      on Press: InvertBit("water_LEVEL_FB")
      Appearance <- "water_LEVEL_FB"
   SymbolLibrary "Symbol library_17" at 664,40 size 58x21
   SymbolLibrary "Symbol library_18" at 480,55 size 41x27
   SymbolLibrary "Symbol library_19" at 482,6 size 44x21
   SymbolLibrary "Symbol library_20" at 750,40 size 31x18
   SymbolLibrary "Symbol library_21" at 327,73 size 65x44
   IOField "I/O field_8" at 339,136 size 87x37; FormatPattern 9999
      ProcessValue <- "HMI_Temperature"
   IOField "I/O field_9" at 339,179 size 87x37; FormatPattern 9999
      ProcessValue <- "HMI_Pressure"
   TextField "Text field_13" at 374,122 size 28x23; Text '*C'
   TextField "Text field_14" at 366,204 size 36x23; Text 'Bar'
   GraphicView "Graphic view_3" at 696,366 size 58x46; Picture "Graphic_10"
   GraphicView "Graphic view_5" at 725,304 size 53x40; Picture "Graphic_11"
   Button "Button_2" at 729,309 size 45x31; TextOff 'Text'
      on Press: ActivateScreen("Alarms", 0)
   TextField "Text field_15" at 366,404 size 45x16; Text 'START'
   TextField "Text field_16" at 444,404 size 37x16; Text 'STOP'
   Button "Button_7" at 695,364 size 60x47; TextOff 'Text'
      on Press: SetBit("HMI_Discharge_Ready_OK")
      on Release: ResetBit("HMI_Discharge_Ready_OK")
   TextField "Text field_17" at 719,398 size 12x16; Text 'Text'
   Button "Button_6" at 270,362 size 56x58; TextOff 'Text'; PictureOff "3bd8051b-cacb-467e-ae66-871dfb0f831b_removalai_preview"
      on Press: SetBit("HMI_Emergency_Stop")
      on Release: ResetBit("HMI_Emergency_Stop")
   SymbolLibrary "V5" at 251,295 size 57x44
      on Activate: function_efd93a16("Water control valve", 0, 0, -1, 0, 1)
      Appearance <- "HMI_V5_Open"
   SymbolLibrary "V6" at 716,17 size 57x44
      on Activate: function_efd93a16("Steam Valve", 0, 0, -1, -1, 1)
      Appearance <- "HMI_V6_Open"
   SymbolLibrary "V8" at 286,51 size 57x44
      ProcessValue <- "HMI_V8_Open"
      Appearance <- "HMI_V8_Open"
      on Press: function_efd93a16("Vacuum valve", 0, 0, -1, -1, 1)
   Button "HmiScreenItemData_1" at 138,366 size 123x46; TextOff 'Reports'; TextOn 'Heating Loop Function'; PictureOff "Navigates to Heating Loop Function for TP700 Comfort 17.0.0.0"; PictureOn "Navigates to Heating Loop Function for TP700 Comfort 17.0.0.0"
      on Press: function_fd03fc5c("Report_1")
   ScreenModuleView "Faceplate_1_1" at 465,17 size 57x44; ScreenModuleType ""
   Switch "Toggle_Horizontal_G" at 608,366 size 80x54; CaptionText 'Switch'; TextOff '0'; TextOn '1'; PictureOn "Toggle_Horizontal_G_On_256c"; PictureOff "Toggle_Horizontal_G_Off_256c"
      ProcessValue <- "HMI_RawMaterial_OK"
   Button "D3_Pushbutton_Pressed_Off_Green" at 355,363 size 70x43; TextOff 'Text'; PictureOff "Design_3_Button_Green_Released_On"; PictureOn "Design_3_Button_Green_Pressed_Off"
      on Press: InvertBit("DB_Process_HMI_Start_Production")
   GraphicIOField "D3_Pilotlight_Red" at 710,122 size 59x46; PictureOff "Design_3_PilotLight_Red_Off"; PictureOn "Design_3_PilotLight_Red_On"
      ProcessValue <- "Red light HMI"
   Button "D3_Pushbutton_Pressed_Off_Red" at 430,362 size 65x46; TextOff 'Text'; PictureOff "Design_3_Button_Red_Released_Off"; PictureOn "Design_3_Button_Red_Pressed_On"
      on Press: SetBit("HMI_Stop_Production")
      on Release: ResetBit("HMI_Stop_Production")
   GraphicIOField "D3_Pilotlight_Green" at 711,175 size 58x44; PictureOff "Design_3_PilotLight_Green_Off"; PictureOn "Design_3_PilotLight_Green_On"
      ProcessValue <- "Green_Light HMI"
   GraphicIOField "D3_Pilotlight_Yellow" at 711,75 size 58x44; PictureOff "Design_3_PilotLight_Yellow_Off"; PictureOn "Design_3_PilotLight_Yellow_On"
      ProcessValue <- "Yellow Light HMI"
   TextField "Text field_12" at 603,341 size 101x20; Text 'Confirm_Raw'
   TextField "Text field_18" at 554,179 size 25x23; Text '%'
   Button "Button_3" at 717,228 size 56x58; TextOff 'Text'; PictureOff "3bd8051b-cacb-467e-ae66-871dfb0f831b_removalai_preview"
      on Press: SetBit("HMI_Reset_System")
      on Release: ResetBit("HMI_Reset_System")
   Button "Button_5" at 720,235 size 57x42; TextOff 'Text'; PictureOn "b967b886-de49-44f2-a9d2-87631f730f4c_removalai_preview"; PictureOff "c8212903-3115-4548-90d4-cb1ba5b5bec7_removalai_preview"
      on Press: SetBit("HMI_Reset_System")
      on Release: ResetBit("HMI_Reset_System")
   SymbolLibrary "Symbol library_4" at 683,89 size 23x202
      on Press: InvertBit("HMI_Door_Locked")
      Visibility <- "HMI_Door_Locked"
   Switch "Lever_Horizontal_1_Mono" at 15,154 size 67x50; CaptionText 'Switch'; TextOff '0'; TextOn '1'; PictureOn "Lever_Horizontal_1_On_mono"; PictureOff "Lever_Horizontal_1_Off_mono"
      on Change: InvertBit("HMI_Manhole_Closed"); InvertBit("Manhole_open_FB")
      ProcessValue <- "Manhole_open_FB"
   TextField "Text field_5" at 2,219 size 21x16; Text 'V1'
   TextField "Text field_8" at 40,219 size 21x16; Text 'V2'
   TextField "Text field_9" at 0,246 size 21x16; Text 'V3'
   TextField "Text field_19" at 37,246 size 21x16; Text 'V4'
   TextField "Text field_20" at 0,275 size 21x16; Text 'V5'
   TextField "Text field_21" at 37,275 size 21x16; Text 'V6'
   TextField "Text field_22" at 0,303 size 21x16; Text 'V7'
   TextField "Text field_23" at 37,303 size 21x16; Text 'V8'
   TextField "Text field_25" at 13,337 size 21x16; Text 'V9'
   GraphicIOField "PlotLight_Round_G" at 18,214 size 22x24; PictureOff "PilotLight_Round_G_Off_256c"; PictureOn "PilotLight_Round_G_On_256c"
      ProcessValue <- "HMI_V1_Open"
   GraphicIOField "PlotLight_Round_G_1" at 18,242 size 22x24; PictureOff "PilotLight_Round_G_Off_256c"; PictureOn "PilotLight_Round_G_On_256c"
      ProcessValue <- "HMI_V3_close"
   GraphicIOField "PlotLight_Round_G_2" at 56,216 size 22x24; PictureOff "PilotLight_Round_G_Off_256c"; PictureOn "PilotLight_Round_G_On_256c"
      ProcessValue <- "HMI_V2_Open"
   GraphicIOField "PlotLight_Round_G_3" at 18,300 size 22x24; PictureOff "PilotLight_Round_G_Off_256c"; PictureOn "PilotLight_Round_G_On_256c"
      ProcessValue <- "HMI_V7_Open"
   GraphicIOField "PlotLight_Round_G_4" at 18,270 size 22x24; PictureOff "PilotLight_Round_G_Off_256c"; PictureOn "PilotLight_Round_G_On_256c"
      ProcessValue <- "HMI_V5_Open"
   GraphicIOField "PlotLight_Round_G_5" at 56,242 size 22x24; PictureOff "PilotLight_Round_G_Off_256c"; PictureOn "PilotLight_Round_G_On_256c"
      ProcessValue <- "HMI_V4_Open"
   GraphicIOField "PlotLight_Round_G_6" at 56,270 size 22x24; PictureOff "PilotLight_Round_G_Off_256c"; PictureOn "PilotLight_Round_G_On_256c"
      ProcessValue <- "HMI_V6_Open"
   GraphicIOField "PlotLight_Round_G_7" at 56,300 size 22x24; PictureOff "PilotLight_Round_G_Off_256c"; PictureOn "PilotLight_Round_G_On_256c"
      ProcessValue <- "HMI_V8_Open"
   GraphicIOField "PlotLight_Round_G_8" at 36,330 size 22x24; PictureOff "PilotLight_Round_G_Off_256c"; PictureOn "PilotLight_Round_G_On_256c"
      ProcessValue <- "HMI_V9_Open"
   Bar "Bar_1" at 152,115 size 31x174; MinimumValue 0; MaximumValue 100
      ProcessValue <- "HMI_Progress"
   Switch "Toggle_Horizontal_G_1" at 519,366 size 80x54; CaptionText 'Switch'; TextOff '0'; TextOn '1'; PictureOn "Toggle_Horizontal_G_On_256c"; PictureOff "Toggle_Horizontal_G_Off_256c"
      ProcessValue <- "HMI_Discharge_Ready_OK"
   TextField "Text field_24" at 510,342 size 92x20; Text 'Confirm_Dis'
   Bar "Bar_2" at 465,268 size 87x64; MinimumValue 0; MaximumValue 100
      ProcessValue <- "Water_level"
      MaximumValue <- "Water Quant."
   GraphicIOField "PlotLight_Round_G_9" at 18,215 size 22x24; PictureOff "PilotLight_Round_G_Off_256c"; PictureOn "Design_3_PilotLight_Red_On"
      ProcessValue <- "HMI_V1_Closed"
   Button "Button_4" at 94,247 size 47x34; TextOff 'Text'; PictureOn "b967b886-de49-44f2-a9d2-87631f730f4c_removalai_preview"; PictureOff "c8212903-3115-4548-90d4-cb1ba5b5bec7_removalai_preview"
      on Press: SetBit("Reset_p_s")
      on Release: ResetBit("Reset_p_s")
   TextField "Text field_26" at 715,280 size 72x23; Text 'Full sys'
   TextField "Text field_27" at 86,225 size 72x23; Text 'Sub sys'
   SymbolLibrary "Symbol library_7" at 185,94 size 8x272
   SymbolLibrary "Symbol library_8" at 187,0 size 8x54
   SymbolLibrary "Symbol library_22" at 780,2 size 20x418
   SymbolLibrary "Symbol library_23" at 457,209 size 34x29
      Appearance <- "Direction Motor"
   SymbolLibrary "Symbol library_24" at 519,209 size 41x31
      Appearance <- "Direction Motor"
   IOField "I/O field_5" at 0,60 size 185x36; FormatPattern ????????????????????????????????????????
      ProcessValue <- "HMI_Status_Message"

screen "Alarms" 800x420, template "Template_1"
   AlarmView "Alarm view_1" at 36,12 size 740x332
   Button "Button_1" at 328,362 size 96x32; TextOff 'Text'
      on Press: function_efd93a16()

PopupScreen "ManHole Valve" 240x240
   TextField "Text field_15" at 45,186 size 45x16; Text 'START'
   Button "Button_3" at 34,138 size 59x45; TextOff 'Text'
      on Press: InvertBit("HMI_V1_Manual_Open")
      Visibility <- "HMI_Process_Running"
   GraphicView "Graphic view_2" at 51,146 size 29x28; Picture "Graphic_12"
   TextField "Text field_16" at 159,185 size 37x16; Text 'STOP'
   Button "Button_4" at 146,138 size 57x44; TextOff 'Text'; PictureOff "Graphic_13"
      on Press: InvertBit("HMI_V1_Manual_Close")
      Visibility <- "HMI_Process_Running"
   TextField "Text field_1" at 13,9 size 224x18; Text 'V1 - MANHOLE VALVE CONTROL'
   SymbolLibrary "Symbol library_7" at 21,43 size 110x73
      ProcessValue <- "HMI_V8_Open"
      Visibility <- "HMI_V1_Open"
   Button "Button_1" at 100,203 size 41x32; TextOff 'Text'; PictureOff "Navigates to Sub Open/Close Manhole for TP700 Comfort 17.0.0.0"
      on Press: ActivateScreen("MAIN LAYOUT SCREEN", 0)
   SymbolLibrary "Symbol library_1" at 126,45 size 110x73
      ProcessValue <- "HMI_V8_Open"
      Visibility <- "HMI_V1_Closed"

PopupScreen "CIP" 240x240
   TextField "Text field_15" at 45,186 size 45x16; Text 'START'
   Button "Button_3" at 34,138 size 59x45; TextOff 'Text'
      on Press: InvertBit("HMI_V2_Manual_Open")
      Visibility <- "HMI_Process_Running"
   GraphicView "Graphic view_2" at 51,146 size 29x28; Picture "Graphic_12"
   TextField "Text field_16" at 159,185 size 37x16; Text 'STOP'
   Button "Button_4" at 146,138 size 57x44; TextOff 'Text'; PictureOff "Graphic_13"
      on Press: InvertBit("HMI_V2_Manual_Close")
      Visibility <- "HMI_Process_Running"
   TextField "Text field_1" at 46,8 size 181x18; Text 'V2 - CIP VALVE CONTROL'
   SymbolLibrary "Symbol library_7" at 21,43 size 110x73
      ProcessValue <- "HMI_V8_Open"
      Visibility <- "HMI_V2_Open"
   Button "Button_1" at 100,203 size 41x32; TextOff 'Text'; PictureOff "Navigates to Sub Open/Close Manhole for TP700 Comfort 17.0.0.0"
      on Press: ActivateScreen("MAIN LAYOUT SCREEN", 0)
   SymbolLibrary "Symbol library_1" at 126,45 size 110x73
      ProcessValue <- "HMI_V8_Open"
      Visibility <- "HMI_V1_Closed"

PopupScreen "Discharge Unlock Valve" 240x240
   TextField "Text field_15" at 45,186 size 45x16; Text 'START'
   Button "Button_3" at 34,138 size 59x45; TextOff 'Text'
      on Press: InvertBit("HMI_V3_Manual_Open")
      Visibility <- "HMI_Process_Running"
   GraphicView "Graphic view_2" at 51,146 size 29x28; Picture "Graphic_12"
   TextField "Text field_16" at 159,185 size 37x16; Text 'STOP'
   Button "Button_4" at 146,138 size 57x44; TextOff 'Text'; PictureOff "Graphic_13"
      on Press: InvertBit("HMI_V3_Manual_Close")
      Visibility <- "HMI_Process_Running"
   TextField "Text field_1" at -8,7 size 248x18; Text 'V3 - DISCHARGE UNLOCK CONTROL'
   SymbolLibrary "Symbol library_7" at 21,43 size 110x73
      ProcessValue <- "HMI_V8_Open"
      Visibility <- "HMI_V3_Open"
   Button "Button_1" at 100,203 size 41x32; TextOff 'Text'; PictureOff "Navigates to Sub Open/Close Manhole for TP700 Comfort 17.0.0.0"
      on Press: ActivateScreen("MAIN LAYOUT SCREEN", 0)
   SymbolLibrary "Symbol library_1" at 126,45 size 110x73
      ProcessValue <- "HMI_V8_Open"
      Visibility <- "HMI_V3_Open"

PopupScreen "Discharge Open" 240x240
   TextField "Text field_15" at 45,186 size 45x16; Text 'START'
   Button "Button_3" at 34,138 size 59x45; TextOff 'Text'
      on Press: InvertBit("HMI_V4_Manual_Open")
      Visibility <- "HMI_Process_Running"
   GraphicView "Graphic view_2" at 51,146 size 29x28; Picture "Graphic_12"
   TextField "Text field_16" at 159,185 size 37x16; Text 'STOP'
   Button "Button_4" at 146,138 size 57x44; TextOff 'Text'; PictureOff "Graphic_13"
      on Press: InvertBit("HMI_V4_Manual_Close")
      Visibility <- "HMI_Process_Running"
   TextField "Text field_1" at 13,9 size 243x18; Text 'V4: "DISCHARGE OPEN CONTROL"'
   SymbolLibrary "Symbol library_7" at 21,43 size 110x73
      ProcessValue <- "HMI_V8_Open"
      Visibility <- "HMI_V4_Open"
   Button "Button_1" at 100,203 size 41x32; TextOff 'Text'; PictureOff "Navigates to Sub Open/Close Manhole for TP700 Comfort 17.0.0.0"
      on Press: ActivateScreen("MAIN LAYOUT SCREEN", 0)
   SymbolLibrary "Symbol library_1" at 126,45 size 110x73
      ProcessValue <- "HMI_V8_Open"
      Visibility <- "HMI_V4_Open"

PopupScreen "Water control valve" 240x240
   TextField "Text field_15" at 45,186 size 45x16; Text 'START'
   GraphicView "Graphic view_2" at 51,146 size 29x28; Picture "Graphic_12"
   TextField "Text field_16" at 159,185 size 37x16; Text 'STOP'
   TextField "Text field_1" at 13,9 size 222x18; Text 'V5: "WATER SUPPLY CONTROL"'
   SymbolLibrary "Symbol library_7" at 21,43 size 106x73
      ProcessValue <- "HMI_V8_Open"
      Appearance <- "HMI_V5_Manual_Open"
   Button "Button_1" at 100,203 size 41x32; TextOff 'Text'; PictureOff "Navigates to Sub Open/Close Manhole for TP700 Comfort 17.0.0.0"
      on Press: ActivateScreen("MAIN LAYOUT SCREEN", 0)
   Button "D3_Pushbutton_Pressed_Off_Green" at 30,142 size 70x43; TextOff 'Text'; PictureOff "Design_3_Button_Green_Released_On"; PictureOn "Design_3_Button_Green_Pressed_Off"
      on Press: InvertBit("HMI_V5_Manual_Open")
   Button "D3_Pushbutton_Pressed_Off_Red" at 141,139 size 65x46; TextOff 'Text'; PictureOff "Design_3_Button_Red_Released_Off"; PictureOn "Design_3_Button_Red_Pressed_On"
      on Press: SetBit("HMI_V5_Manual_Close")
   SymbolLibrary "Symbol library_2" at 127,43 size 106x73
      ProcessValue <- "HMI_V8_Open"
      Appearance <- "HMI_V5_Manual_Close"

PopupScreen "Steam Valve" 240x240
   TextField "Text field_1" at 13,9 size 217x18; Text 'V6: "STEAM VALVE CONTROL"'
   Button "Button_1" at 100,203 size 41x32; TextOff 'Text'; PictureOff "Navigates to Sub Open/Close Manhole for TP700 Comfort 17.0.0.0"
      on Press: ActivateScreen("MAIN LAYOUT SCREEN", 0)
   TextField "Text field_15" at 45,186 size 45x16; Text 'START'
   TextField "Text field_16" at 159,185 size 37x16; Text 'STOP'
   SymbolLibrary "Symbol library_7" at 21,43 size 106x73
      ProcessValue <- "HMI_V8_Open"
      Appearance <- "HMI_V6_Manual_Open"
   Button "D3_Pushbutton_Pressed_Off_Green" at 30,142 size 70x43; TextOff 'Text'; PictureOff "Design_3_Button_Green_Released_On"; PictureOn "Design_3_Button_Green_Pressed_Off"
      on Press: InvertBit("HMI_V6_Manual_Open")
   Button "D3_Pushbutton_Pressed_Off_Red" at 141,139 size 65x46; TextOff 'Text'; PictureOff "Design_3_Button_Red_Released_Off"; PictureOn "Design_3_Button_Red_Pressed_On"
      on Press: SetBit("HMI_V6_Manual_Close")
   SymbolLibrary "Symbol library_2" at 127,43 size 106x73
      ProcessValue <- "HMI_V8_Open"
      Appearance <- "HMI_V6_Manual_Close"

PopupScreen "Evacuation valve" 240x240
   TextField "Text field_15" at 45,186 size 45x16; Text 'START'
   Button "Button_3" at 34,138 size 59x45; TextOff 'Text'
      on Press: InvertBit("HMI_V7_Manual_Open")
      Visibility <- "HMI_Process_Running"
   GraphicView "Graphic view_2" at 51,146 size 29x28; Picture "Graphic_12"
   TextField "Text field_16" at 159,185 size 37x16; Text 'STOP'
   Button "Button_4" at 146,138 size 57x44; TextOff 'Text'; PictureOff "Graphic_13"
      on Press: InvertBit("HMI_V7_Manual_Close")
      Visibility <- "HMI_Process_Running"
   TextField "Text field_1" at 9,32 size 231x16; Text 'V7: "EVACUATION VALVE CONTROL"'
   SymbolLibrary "Symbol library_7" at 20,59 size 110x73
      ProcessValue <- "HMI_V8_Open"
      Visibility <- "HMI_V7_Open"
   Button "Button_1" at 100,203 size 41x32; TextOff 'Text'; PictureOff "Navigates to Sub Open/Close Manhole for TP700 Comfort 17.0.0.0"
      on Press: ActivateScreen("MAIN LAYOUT SCREEN", 0)
   SymbolLibrary "Symbol library_1" at 127,59 size 110x73
      ProcessValue <- "HMI_V8_Open"
      Visibility <- "HMI_V7_Open"

PopupScreen "Vacuum valve" 240x240
   TextField "Text field_1" at 13,9 size 223x18; Text 'V8: "VACUUM VALVE CONTROL"'
   SymbolLibrary "Symbol library_7" at 21,43 size 110x73
      ProcessValue <- "HMI_V8_Open"
      Appearance <- "HMI_V8_Manual_Open"
      Visibility <- "HMI_V8_Manual_Close"
   Button "Button_1" at 100,203 size 41x32; TextOff 'Text'; PictureOff "Navigates to Sub Open/Close Manhole for TP700 Comfort 17.0.0.0"
      on Press: ActivateScreen("MAIN LAYOUT SCREEN", 0)
   SymbolLibrary "Symbol library_1" at 126,45 size 110x73
      ProcessValue <- "HMI_V8_Open"
      Visibility <- "HMI_V8_Manual_Open"
      Appearance <- "HMI_V8_Manual_Close"
   TextField "Text field_15" at 45,185 size 45x16; Text 'START'
   TextField "Text field_16" at 159,185 size 37x16; Text 'STOP'
   SymbolLibrary "Symbol library_2" at 21,43 size 106x73
      ProcessValue <- "HMI_V8_Open"
      Appearance <- "HMI_V8_Manual_Open"
   Button "D3_Pushbutton_Pressed_Off_Green_1" at 30,142 size 70x43; TextOff 'Text'; PictureOff "Design_3_Button_Green_Released_On"; PictureOn "Design_3_Button_Green_Pressed_Off"
      on Press: InvertBit("HMI_V8_Manual_Open")
   Button "D3_Pushbutton_Pressed_Off_Red_1" at 141,139 size 65x46; TextOff 'Text'; PictureOff "Design_3_Button_Red_Released_Off"; PictureOn "Design_3_Button_Red_Pressed_On"
      on Press: SetBit("HMI_V8_Manual_Close")
   SymbolLibrary "Symbol library_3" at 127,43 size 106x73
      ProcessValue <- "HMI_V8_Open"
      Appearance <- "HMI_V8_Manual_Close"

PopupScreen "Vacuum cooling" 240x240
   TextField "Text field_15" at 45,186 size 45x16; Text 'START'
   Button "Button_3" at 34,138 size 59x45; TextOff 'Text'
      on Press: InvertBit("HMI_V9_Manual_Open")
      Visibility <- "HMI_Process_Running"
   GraphicView "Graphic view_2" at 51,146 size 29x28; Picture "Graphic_12"
   TextField "Text field_16" at 159,185 size 37x16; Text 'STOP'
   Button "Button_4" at 146,138 size 57x44; TextOff 'Text'; PictureOff "Graphic_13"
      on Press: InvertBit("HMI_V9_Manual_Close")
      Visibility <- "HMI_Process_Running"
   TextField "Text field_1" at 13,9 size 240x18; Text 'V9: "VACUUM COOLING CONTROL"'
   SymbolLibrary "Symbol library_7" at 21,43 size 110x73
      ProcessValue <- "HMI_V8_Open"
      Visibility <- "HMI_V9_Open"
   Button "Button_1" at 100,203 size 41x32; TextOff 'Text'; PictureOff "Navigates to Sub Open/Close Manhole for TP700 Comfort 17.0.0.0"
      on Press: ActivateScreen("MAIN LAYOUT SCREEN", 0)
   SymbolLibrary "Symbol library_1" at 126,45 size 110x73
      ProcessValue <- "HMI_V8_Open"
      Visibility <- "HMI_V9_Open"

PopupScreen "motor manual" 240x240
   TextField "Text field_15" at 45,186 size 45x16; Text 'START'
   Button "Button_3" at 34,138 size 59x45; TextOff 'Text'
      on Press: InvertBit("HMI_V6_Manual_Open")
      Visibility <- "HMI_Process_Running"
   GraphicView "Graphic view_2" at 51,146 size 29x28; Picture "Graphic_12"
   TextField "Text field_16" at 122,184 size 37x16; Text 'STOP'
   Button "Button_4" at 111,142 size 57x44; TextOff 'Text'; PictureOff "Graphic_13"
      on Press: InvertBit("HMI_V6_Manual_Close")
      Visibility <- "HMI_Process_Running"
   Button "Button_1" at 81,206 size 41x32; TextOff 'Text'; PictureOff "Navigates to Sub Open/Close Manhole for TP700 Comfort 17.0.0.0"
      on Press: ActivateScreen("MAIN LAYOUT SCREEN", 0)
   SymbolLibrary "Symbol library_1" at 12,6 size 104x70
   SymbolicIOField "Symbolic I/O field_1" at 34,98 size 86x27; TextOff '0'; TextOn '1'
      ProcessValue <- "HMI_Motor_Speed"
   Gauge "Gauge_1" at 145,11 size 114x114; CaptionText 'Speed'; UnitText 'rpm'
      ProcessValue <- "HMI_Motor_Speed"
      MaximumValue <- "DB_Motors_Motors{1}_Config_Max_Speed_pct"
      MinimumValue <- "DB_Motors_Motors{1}_Config_Min_Speed_pct"

PopupScreen "parameters" 240x240
   IOField "I/O field_1" at 129,0 size 96x32; FormatPattern 999
      ProcessValue <- "Cooking Time"
   TextField "Text field_1" at 0,0 size 129x23; Text 'Cooking Time'
   IOField "I/O field_2" at 129,32 size 96x32; FormatPattern 999
      ProcessValue <- "Cold Mix Time"
   TextField "Text field_3" at 0,32 size 134x23; Text 'Cold Mix Time'
   IOField "I/O field_3" at 129,64 size 96x32; FormatPattern s999999999.999
      ProcessValue <- "Water Quant."
   TextField "Text field_5" at 0,64 size 142x23; Text 'Water quantity'
   TextField "Text field_6" at 225,64 size 15x23; Text 'L'
   IOField "I/O field_4" at 126,91 size 96x32; FormatPattern s9999999999
      ProcessValue <- "Forward Time"
   TextField "Text field_7" at 0,96 size 130x23; Text 'Forward Time'
   IOField "I/O field_5" at 125,124 size 96x32; FormatPattern s9999999999
      ProcessValue <- "FB_Motor_VFD_DB_Tmr_Bwd_PT"
   TextField "Text field_9" at 0,124 size 144x23; Text 'Backward Time'
   IOField "I/O field_6" at 125,155 size 96x32; FormatPattern s999999999.999
      ProcessValue <- "Water Quant."
   TextField "Text field_11" at 0,160 size 117x23; Text 'Vacuum Set.'

PopupScreen "Vacuum valve_1" 240x240
   TextField "Text field_1" at 13,9 size 223x18; Text 'V8: "VACUUM VALVE CONTROL"'
   SymbolLibrary "Symbol library_7" at 21,43 size 110x73
      ProcessValue <- "HMI_V8_Open"
      Appearance <- "HMI_V8_Manual_Open"
      Visibility <- "HMI_V8_Manual_Close"
   Button "Button_1" at 100,203 size 41x32; TextOff 'Text'; PictureOff "Navigates to Sub Open/Close Manhole for TP700 Comfort 17.0.0.0"
      on Press: ActivateScreen("MAIN LAYOUT SCREEN", 0)
   SymbolLibrary "Symbol library_1" at 126,45 size 110x73
      ProcessValue <- "HMI_V8_Open"
      Visibility <- "HMI_V8_Manual_Open"
      Appearance <- "HMI_V8_Manual_Close"
   Button "D3_Pushbutton_Pressed_Off_Red" at 125,136 size 65x46; TextOff 'Text'; PictureOff "Design_3_Button_Red_Released_Off"; PictureOn "Design_3_Button_Red_Pressed_On"
      on Press: SetBit("HMI_V8_Manual_Close")
      on Release: ResetBit("HMI_V8_Manual_Close")
   TextField "Text field_2" at 61,178 size 45x16; Text 'START'
   TextField "Text field_3" at 139,178 size 37x16; Text 'STOP'
   Button "D3_Pushbutton_Pressed_Off_Green" at 50,137 size 70x43; TextOff 'Text'; PictureOff "Design_3_Button_Green_Released_On"; PictureOn "Design_3_Button_Green_Pressed_Off"
      on Press: InvertBit("HMI_V8_Manual_Open")

PopupScreen "Vacuum valve_2" 240x240
   TextField "Text field_1" at 13,9 size 223x18; Text 'V8: "VACUUM VALVE CONTROL"'
   SymbolLibrary "Symbol library_7" at 21,43 size 110x73
      ProcessValue <- "HMI_V8_Open"
      Appearance <- "HMI_V8_Manual_Open"
      Visibility <- "HMI_V8_Manual_Close"
   Button "Button_1" at 100,203 size 41x32; TextOff 'Text'; PictureOff "Navigates to Sub Open/Close Manhole for TP700 Comfort 17.0.0.0"
      on Press: ActivateScreen("MAIN LAYOUT SCREEN", 0)
   SymbolLibrary "Symbol library_1" at 126,45 size 110x73
      ProcessValue <- "HMI_V8_Open"
      Visibility <- "HMI_V8_Manual_Open"
      Appearance <- "HMI_V8_Manual_Close"
   Button "D3_Pushbutton_Pressed_Off_Red" at 125,136 size 65x46; TextOff 'Text'; PictureOff "Design_3_Button_Red_Released_Off"; PictureOn "Design_3_Button_Red_Pressed_On"
      on Press: SetBit("HMI_V8_Manual_Close")
      on Release: ResetBit("HMI_V8_Manual_Close")
   TextField "Text field_2" at 61,178 size 45x16; Text 'START'
   TextField "Text field_3" at 139,178 size 37x16; Text 'STOP'
   Button "D3_Pushbutton_Pressed_Off_Green" at 50,137 size 70x43; TextOff 'Text'; PictureOff "Design_3_Button_Green_Released_On"; PictureOn "Design_3_Button_Green_Pressed_Off"
      on Press: InvertBit("HMI_V8_Manual_Open")
*)

(* ===== HMI "HMI_RT_1" =====

ScreenModuleEditorView "Faceplate_1" 640x480
   SymbolLibrary "V7" at 10,10 size 57x44
*)

(* ===== HMI "HMI_RT_1" =====

ScreenModuleEditorView "Faceplate_1" 640x480
   SymbolLibrary "V7" at 126,24 size 57x44
*)

(* ===== HMI "HMI_RT_1" =====

ScreenModuleEditorView "Faceplate_1" 640x480
   SymbolLibrary "V7" at 10,10 size 57x44
*)